ABB RAPID module: SpeedProg.mod

%%%
  VERSION:1
  LANGUAGE:ENGLISH
%%%
MODULE MOD_SpeedProg

    ! -------------------------------
    ! Define customized variables here
    ! ...

	! Tool variables:
	PERS tooldata ToolS := [TRUE,[[10.000,20.000,150.000],[1.00000000,0.00000000,0.00000000,0.00000000]],[1,[0,0,20],[1,0,0,0],0,0,0.005]];

	! Reference variables:
	PERS wobjdata FrameS := [FALSE, TRUE, "", [[0,0,0],[1,0,0,0]],[[1234.570,-98.765,50.500],[0.96592583,0.00000000,0.00000000,0.25881905]]];

	PROC Main()
		ConfJ \On;
		ConfL \Off;
		! Program generated by RoboDK v6.0.7 for ABB IRBT 2005 Standard 2.8m on XX/XX/XXXX 18:00:00
		! Using nominal kinematics.
		MoveL [[-607.850,543.849,363.215],[0.37410804,0.28584607,0.85365954,-0.22271191],[0,0,0,0],[9E+09,9E+09,9E+09,9E+09,9E+09,9E+09]],[1.00,500,5000,1000],[FALSE,0.3,0.4,0.4,0.0,0.4,0.0],ToolS \WObj:=FrameS;
		MoveAbsJ [[250.000000,0.000000,0.000000,0.000000,0.000000,0.000000],[9E+09,9E+09,9E+09,9E+09,9E+09,9E+09]],[1.00,500,5000,1000],[FALSE,0.3,0.4,0.4,0.0,0.4,0.0],ToolS \WObj:=FrameS;
		MoveL [[-640.584,506.980,371.534],[0.37410804,0.28584607,0.85365954,-0.22271191],[0,0,0,0],[9E+09,9E+09,9E+09,9E+09,9E+09,9E+09]],[12.30,500,5000,1000],z1,ToolS \WObj:=FrameS;
		MoveAbsJ [[500.000000,0.000000,0.000000,0.000000,0.000000,0.000000],[9E+09,9E+09,9E+09,9E+09,9E+09,9E+09]],[12.30,500,5000,1000],z1,ToolS \WObj:=FrameS;
		MoveL [[-607.850,543.849,363.215],[0.37410804,0.28584607,0.85365954,-0.22271191],[0,0,0,0],[9E+09,9E+09,9E+09,9E+09,9E+09,9E+09]],[99.90,500,5000,1000],[FALSE,2.5,3.8,3.8,0.4,3.8,0.4],ToolS \WObj:=FrameS;
		MoveAbsJ [[250.000000,0.000000,0.000000,0.000000,0.000000,0.000000],[9E+09,9E+09,9E+09,9E+09,9E+09,9E+09]],[99.90,500,5000,1000],[FALSE,2.5,3.8,3.8,0.4,3.8,0.4],ToolS \WObj:=FrameS;
		MoveL [[-640.584,506.980,371.534],[0.37410804,0.28584607,0.85365954,-0.22271191],[0,0,0,0],[9E+09,9E+09,9E+09,9E+09,9E+09,9E+09]],[333.33,500,5000,1000],[FALSE,3.7,5.6,5.6,0.6,5.6,0.6],ToolS \WObj:=FrameS;
		MoveAbsJ [[500.000000,0.000000,0.000000,0.000000,0.000000,0.000000],[9E+09,9E+09,9E+09,9E+09,9E+09,9E+09]],[333.33,500,5000,1000],[FALSE,3.7,5.6,5.6,0.6,5.6,0.6],ToolS \WObj:=FrameS;
		MoveL [[-607.850,543.849,363.215],[0.37410804,0.28584607,0.85365954,-0.22271191],[0,0,0,0],[9E+09,9E+09,9E+09,9E+09,9E+09,9E+09]],v1000,[FALSE,6.0,9.0,9.0,0.9,9.0,0.9],ToolS \WObj:=FrameS;
		MoveAbsJ [[250.000000,0.000000,0.000000,0.000000,0.000000,0.000000],[9E+09,9E+09,9E+09,9E+09,9E+09,9E+09]],v1000,[FALSE,6.0,9.0,9.0,0.9,9.0,0.9],ToolS \WObj:=FrameS;
		MoveL [[-640.584,506.980,371.534],[0.37410804,0.28584607,0.85365954,-0.22271191],[0,0,0,0],[9E+09,9E+09,9E+09,9E+09,9E+09,9E+09]],v2500,[FALSE,9.0,13.5,13.5,1.4,13.5,1.4],ToolS \WObj:=FrameS;
		MoveAbsJ [[500.000000,0.000000,0.000000,0.000000,0.000000,0.000000],[9E+09,9E+09,9E+09,9E+09,9E+09,9E+09]],v2500,[FALSE,9.0,13.5,13.5,1.4,13.5,1.4],ToolS \WObj:=FrameS;
		MoveL [[-607.850,543.849,363.215],[0.37410804,0.28584607,0.85365954,-0.22271191],[0,0,0,0],[9E+09,9E+09,9E+09,9E+09,9E+09,9E+09]],v5000,z15,ToolS \WObj:=FrameS;
		MoveAbsJ [[250.000000,0.000000,0.000000,0.000000,0.000000,0.000000],[9E+09,9E+09,9E+09,9E+09,9E+09,9E+09]],v5000,z15,ToolS \WObj:=FrameS;
		MoveL [[-640.584,506.980,371.534],[0.37410804,0.28584607,0.85365954,-0.22271191],[0,0,0,0],[9E+09,9E+09,9E+09,9E+09,9E+09,9E+09]],v7000,z30,ToolS \WObj:=FrameS;
		MoveAbsJ [[500.000000,0.000000,0.000000,0.000000,0.000000,0.000000],[9E+09,9E+09,9E+09,9E+09,9E+09,9E+09]],v7000,z30,ToolS \WObj:=FrameS;
		MoveL [[-607.850,543.849,363.215],[0.37410804,0.28584607,0.85365954,-0.22271191],[0,0,0,0],[9E+09,9E+09,9E+09,9E+09,9E+09,9E+09]],[0.50,500,5000,1000],[FALSE,75.0,112.5,112.5,11.2,112.5,11.2],ToolS \WObj:=FrameS;
		MoveAbsJ [[250.000000,0.000000,0.000000,0.000000,0.000000,0.000000],[9E+09,9E+09,9E+09,9E+09,9E+09,9E+09]],[0.50,500,5000,1000],[FALSE,75.0,112.5,112.5,11.2,112.5,11.2],ToolS \WObj:=FrameS;
		MoveL [[-640.584,506.980,371.534],[0.37410804,0.28584607,0.85365954,-0.22271191],[0,0,0,0],[9E+09,9E+09,9E+09,9E+09,9E+09,9E+09]],[750.00,500,5000,1000],z150,ToolS \WObj:=FrameS;
		MoveAbsJ [[500.000000,0.000000,0.000000,0.000000,0.000000,0.000000],[9E+09,9E+09,9E+09,9E+09,9E+09,9E+09]],[750.00,500,5000,1000],z150,ToolS \WObj:=FrameS;
		MoveL [[-640.584,506.980,371.534],[0.37410804,0.28584607,0.85365954,-0.22271191],[0,0,0,0],[9E+09,9E+09,9E+09,9E+09,9E+09,9E+09]],[750.00,500,5000,1000],z150,ToolS \WObj:=FrameS;
	ENDPROC

ENDMODULE
